(* IEC 61131-3 sources: plc_generation_empirical_study/datasets/packages/internal_v0_1/qualification_only/C01_E01_two_input_permissive, 1 file *)

(* ---- reference.st ---- *)
FUNCTION_BLOCK C01_E01_two_input_permissive
VAR_INPUT
    Enable : BOOL;
    GuardClosed : BOOL;
END_VAR
VAR_OUTPUT
    RunPermit : BOOL;
END_VAR

RunPermit := Enable AND GuardClosed;

END_FUNCTION_BLOCK
